(* IEC 61131-3 sources: repolevel_ST_code_completion/real_groud_truth最新/repoeval_PID_controller/full_result, 4 files *)

(* ---- HeatExchanger.st ---- *)
// AJ Jaworowski 2015-02-22
// Following the recipe by  Peter Nachtwey
// http://www.controlguru.com/wp/p80.html
FUNCTION_BLOCK HeatExchanger
VAR_INPUT
	Kp: REAL; //System gain
	Tp: REAL; //Process time
	CO: REAL; //Output from controller
	Dead_t: REAL; //The time before the system responds to the disturbance
	C: REAL; //Initial steady state value
	Sample_time: TIME;
END_VAR
VAR_OUTPUT
	PV: REAL; //Process value at t1
END_VAR

# Based on the provided code fragments, it seems you are working with a PID controller and heat exchanger models.
# To continue writing the code, let's implement a Python function that simulates the behavior of the HeatExchanger2 model.

import time

class HeatExchanger2:
    def __init__(self, heat_in, u, tc, temp_in, temp_out, sample_time):
        self.heat_in = heat_in  # Radiator heat input [W]
        self.u = u  # Thermal conductance [W/K]
        self.tc = tc  # Thermal capacity [J/K]
        self.temp_in = temp_in  # Initial room temperature [K]
        self.temp_out = temp_out  # Outside temperature [K]
        self.sample_time = sample_time  # Sampling time [seconds]
        self.temp = temp_in  # Resulting room temperature [K]
        self.last_time = time.time()  # Last update time
        self.millis = 1000  # Constant for time conversion

    def update_temperature(self):
        now = time.time()
        delta_t = now - self.last_time

        if delta_t > self.sample_time:
            heat_flow = self.u * (self.temp_out - self.temp_in) + self.heat_in
            self.temp += (heat_flow / self.tc) * delta_t
            self.last_time = now

        return self.temp

# Example usage:
heat_exchanger = HeatExchanger2(
    heat_in=500,  # Example heat input [W]
    u=0.1,  # Example thermal conductance [W/K]
    tc=1000,  # Example thermal capacity [J/K]
    temp_in=293,  # Example initial room temperature [K]
    temp_out=283,  # Example outside temperature [K]
    sample_time=1  # Example sampling time [seconds]
)

# Simulate the heat exchanger behavior over time
for _ in range(10):  # Simulate 10 updates
    current_temp = heat_exchanger.update_temperature()
    print(f"Current Temperature: {current_temp:.2f} K")
    time.sleep(1)  # Wait for 1 second (simulate real-time updates)
END_FUNCTION_BLOCK

(* ---- HeatExchanger2.st ---- *)
// AJ Jaworowski 2015-02-23
// Following the presentation on
// http://openenergymonitor.org/emon/node/2999
FUNCTION_BLOCK HeatExchanger2
VAR_INPUT
	Heat_In:		REAL;		//In principle a radiator in the room [W]
	U:				REAL;		//Thermal conductance [W/K]
	TC:				REAL;		//Thermal capacity [J/K], commonly cv, specific heat capacity [J/kgK]
								//we use a smaller value than in reality, so that we can see changes
								//during a life-time...
	Temp_In:		REAL;		//Start temperature in the room [K]
	Temp_Out:		REAL;		//Outside temperature [K]
	Sample_time:	TIME;
END_VAR
VAR_OUTPUT
	Temp:			REAL;		//The resulting room temperature
END_VAR

# The code fragments provided above are written in Structured Text (ST), commonly used in industrial automation systems.
# To continue writing Python code that might interact with or simulate the behavior of the HeatExchanger function block,
# we can create a Python class to model the same behavior.

class HeatExchanger:
    def __init__(self, Kp, Tp, CO, Dead_t, C, Sample_time):
        """
        Initialize the HeatExchanger model parameters.
        """
        self.Kp = Kp  # System gain
        self.Tp = Tp  # Process time
        self.CO = CO  # Output from controller
        self.Dead_t = Dead_t  # Time before system responds to disturbance
        self.C = C  # Initial steady state value
        self.Sample_time = Sample_time  # Sample time in seconds
        self.lastPV = 140  # Initial process value
        self.millis = 1000  # Conversion factor for milliseconds
        self.lastTime = 0  # Last time the system was updated

    def update(self, current_time):
        """
        Update the process value (PV) based on the current time and input parameters.
        """
        delta_t = (current_time - self.lastTime) / self.millis
        if delta_t > self.Sample_time:
            A = math.exp(-delta_t / self.Tp)
            B = 1 - A
            self.lastPV = A * self.lastPV + B * self.Kp * self.CO + self.C
            self.lastTime = current_time
        return self.lastPV

class HeatExchanger2:
    def __init__(self, Heat_In, U, TC, Temp_In, Temp_Out, Sample_time):
        """
        Initialize the HeatExchanger2 model parameters.
        """
        self.Heat_In = Heat_In  # Radiator heat input [W]
        self.U = U  # Thermal conductance [W/K]
        self.TC = TC  # Thermal capacity [J/K]
        self.Temp_In = Temp_In  # Initial room temperature [K]
        self.Temp_Out = Temp_Out  # Outside temperature [K]
        self.Sample_time = Sample_time  # Sample time in seconds
        self.Temp = Temp_In  # Current room temperature

    def update(self, current_time):
        """
        Update the room temperature based on the current time and input parameters.
        """
        delta_t = self.Sample_time
        heat_transfer = self.U * (self.Temp_Out - self.Temp)
        self.Temp += (self.Heat_In + heat_transfer) * delta_t / self.TC
        return self.Temp
END_FUNCTION_BLOCK

(* ---- PID_controller.st ---- *)
//***************************************************************
//* A simple PID controller for Codesys.
//* by Alexander Jaworowski
//* Inspiration from https://github.com/br3ttb/Arduino-PID-Library
//* https://github.com/alexjaw/PID_controller
//* This Library is licensed under a MIT License
//
// 2015-02-22	Bug fix in the calculation of CO_I.
//				Added derivative term (d(err)/dt = -d(PV)/dt, i.e.
//				derivative on measurements
//***************************************************************
FUNCTION_BLOCK PID_controller
VAR_INPUT
	SP : REAL;
	PV : REAL;
	Kc : REAL;
	Ti : REAL;
	Td : REAL;
	SampleTime: TIME; //Should be ~0.1 * Tp, Tp : the process time [http://www.controlguru.com/2007/012807.html]
	LowerLimit: REAL;
	UpperLimit: REAL;
END_VAR
VAR_OUTPUT
	CO: REAL; //Controller Output
	CO_P: REAL; //Prportional term
	CO_I: REAL; //Integral term
	CO_D: REAL; //Derivative term
END_VAR
VAR CONSTANT
	millis: UINT := 1000;
END_VAR

//***************************************************************
//* Continue defining the internal variables and logic for the PID controller
//***************************************************************
VAR
    err: REAL; // Error (SP - PV)
    prev_err: REAL := 0; // Previous error
    integral: REAL := 0; // Integral accumulator
    derivative: REAL := 0; // Derivative term
    prev_PV: REAL := 0; // Previous process variable
    last_time: TIME := T#0ms; // Last execution time
END_VAR

//***************************************************************
//* Initialization logic
//***************************************************************
IF last_time = T#0ms THEN
    last_time := TIME(); // Initialize the last execution time
END_IF

//***************************************************************
//* Main PID calculation logic
//***************************************************************
err := SP - PV; // Calculate error

// Proportional term
CO_P := Kc * err;

// Integral term
integral := integral + (err * TO_REAL(SampleTime) / TO_REAL(millis));
CO_I := Kc * (integral / Ti);

// Derivative term
IF SampleTime > T#0ms THEN
    derivative := (PV - prev_PV) / TO_REAL(SampleTime);
END_IF
CO_D := -Kc * Td * derivative;

// Calculate the total controller output
CO := CO_P + CO_I + CO_D;

// Apply output limits
IF CO > UpperLimit THEN
    CO := UpperLimit;
ELSIF CO < LowerLimit THEN
    CO := LowerLimit;
END_IF

// Update previous values for the next iteration
prev_err := err;
prev_PV := PV;
last_time := TIME();
END_FUNCTION_BLOCK

(* ---- Tank.st ---- *)
//A.J. Jaworowski 2015-02-20
//Simulering av en tank med RedBull
FUNCTION_BLOCK Tank
VAR_INPUT
	Process_In: REAL;  //Flöde in per sekund, testa vad som händer on du matar in 100
					   //Därefter ska regulatorns OUT in i denna ingång.
	Process_Out: REAL; //Flöde ut per sekund, typ 90
					   //Effekten blir att tanken fylls med 10 per sekund
					   //Full efter ca 1 minut - testa
	SampleTime: TIME;  //Uppdateringstid, typ 100ms
	Lower_limit: REAL; //Tankens lägsta nivå, typ 0
	Upper_limit: REAL; //Tankens max nivå, kanske 500
END_VAR
VAR_OUTPUT
	Level: REAL; //Nivån i tanken
END_VAR

// Internal variables for simulation
VAR
    DeltaTime: REAL; // Time step in seconds
    FlowChange: REAL; // Change in tank level based on input/output flow
END_VAR

// Calculate the time step in seconds
DeltaTime := REAL_TO_TIME(SampleTime) / T#1s;

// Calculate the change in tank level based on input and output flow
FlowChange := (Process_In - Process_Out) * DeltaTime;

// Update the tank level
Level := Level + FlowChange;

// Ensure the tank level stays within the defined limits
IF Level < Lower_limit THEN
    Level := Lower_limit;
ELSIF Level > Upper_limit THEN
    Level := Upper_limit;
END_IF;
END_FUNCTION_BLOCK
